(* IEC 61131-3 sources: katsuragi/st/test, 3 files *)

(* ---- empty_program.st ---- *)
PROGRAM empty_program
END_PROGRAM

(* ---- empty_program_with_comment.st ---- *)
PROGRAM empty_program_with_comment
// line comment

// line comment
// line comment

/* block comment */

/*
 * block comment
 */

(* block comment *)

(*
 * block comment
 *)
END_PROGRAM

(* ---- variable_assignment.st ---- *)
PROGRAM variable_assignment
VAR
	x : INT;
END_VAR

x := 1;

END_PROGRAM
